// TIA Portal V21 export
// export: Created 2026-11-11T00:47:47.468354Z, ExportSetting WithDefaults, DisplayName Totally Integrated Automation Portal, DisplayVersion V21 Update 3, DisplayName STEP 7 Professional, DisplayVersion V21 Update 3, DisplayName STEP 7 Safety, DisplayVersion V21, DisplayName Tech WebApplication, DisplayVersion V21, DisplayName WinCC Basic/Comfort/Advanced, DisplayVersion V21 Update 3, DisplayName WinCC Unified, DisplayVersion V21 Update 3
FUNCTION_BLOCK "FB_Fbd_sc005"   // FB184, FBD
{ S7_Optimized_Access := 'TRUE' }
VERSION : 0.1
// stored: AutoNumber true, IsIECCheckEnabled false, IsRetainMemResEnabled false, MemoryReserve 100, SetENOAutomatically false, UDAEnableTagReadback false
   VAR_INPUT
      v_req : Bool;
      v_r : Bool;
      v_id : CONN_PRG;
      v_r_id : CONN_R_ID;
   END_VAR
   VAR_OUTPUT
      v_done : Bool;
      v_error : Bool;
      v_status : Word;
   END_VAR
   VAR_IN_OUT
      v_sd_1 : Array[0..99] of Byte;
      v_len : Word;
   END_VAR
   VAR
      inst { S7_SetPoint := 'True'} : BSEND;
   END_VAR
BEGIN

REGION Network 1: BSEND - Send data in segments
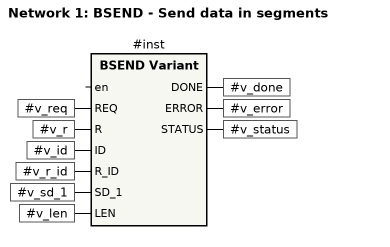
   #inst(REQ := #v_req,   // BSEND
         R := #v_r,
         ID := #v_id,
         R_ID := #v_r_id,
         SD_1 := #v_sd_1,
         LEN := #v_len,
         DONE => #v_done,
         ERROR => #v_error,
         STATUS => #v_status);
END_REGION
END_FUNCTION_BLOCK
